Fanuc KAREL source: KB00079.KL

PROGRAM KB00079
%NOLOCKGROUP
VAR
  P1: INTEGER
  P2: INTEGER
  P3: INTEGER
  RESULT: JOINTPOS
BEGIN
  P1 = 1
  P2 = 1
  P3 = 1
  RESULT = GET_JPOS_TPE(P1, P2, P3)
END KB00079
